(* Schneider Machine Expert - Basic project PROJECT, file version 2.9.0.0 *)
(* ProjectInformations: Name=New project *)

HARDWARE
  Cpu 0: TM221CE16R
  EthernetConfiguration: NetworkName=M221, IpAllocationMode=FixedAddress, IpAddress=0.0.0.0, SubnetMask=0.0.0.0
  SerialLineConfiguration: Baud=Baud19200, Parity=ParityEven, DataBits=DataBits8, StopBits=StopBits1, PhysicalMedium=PhysicalMediumRs485, TransmissionMode=TransmissionModeModbusRtu, SlaveId=1, Addressing=SlaveAddressing
  MastTask: UsePeriodScanMode=false, PeriodScan=100
  FastTask: Period=255
  CpuBehavior: StartingMode=StartAsPreviousState, AutoSaveRamOnEeprom=true, WatchdogPeriod=250

SYMBOLS  (address, symbol, comment, settings)
  %M0         "START"
  %M1         "STOP N RESET"
  %M2         "END CYCLE"
  %M3         "END A"
  %M4         "END B"
  %M10        "BT_START"
  %M11        "BT_RESET"
  %M12        "LAMP IND"
  %M13        "ST VALVE A"
  %M14        "ST VALVE B"
  %M15        "ST VALVE C"
  %M16        "ST AGITATOR"
  %M17        "ST HEATER"
  %M18        "ALARM"
  %S6       SB_TB1S  "Time base of 1 s generated by an internal clock"
  %TM0        "TIMER A"  [Preset=5, Base=OneSecond]
  %TM1        "TIMER B"  [Preset=10, Base=OneSecond]
  %C0         "COUNTER"  [Preset=2]
  %SC0        "COUNTER"
  %I0.0       "START"
  %I0.1       "STOP"
  %I0.2       "SENSOR TINGGI"
  %I0.3       "SENSOR SUHU"
  %Q0.0       "LAMP_INDIKATOR"
  %Q0.1       "VALVE A"
  %Q0.2       "VALVE B"
  %Q0.3       "AGITATOR"
  %Q0.4       "HEATER"
  %Q0.5       "DRAIN VALVE"

POU New POU
  (* SectionNumber=1 *)

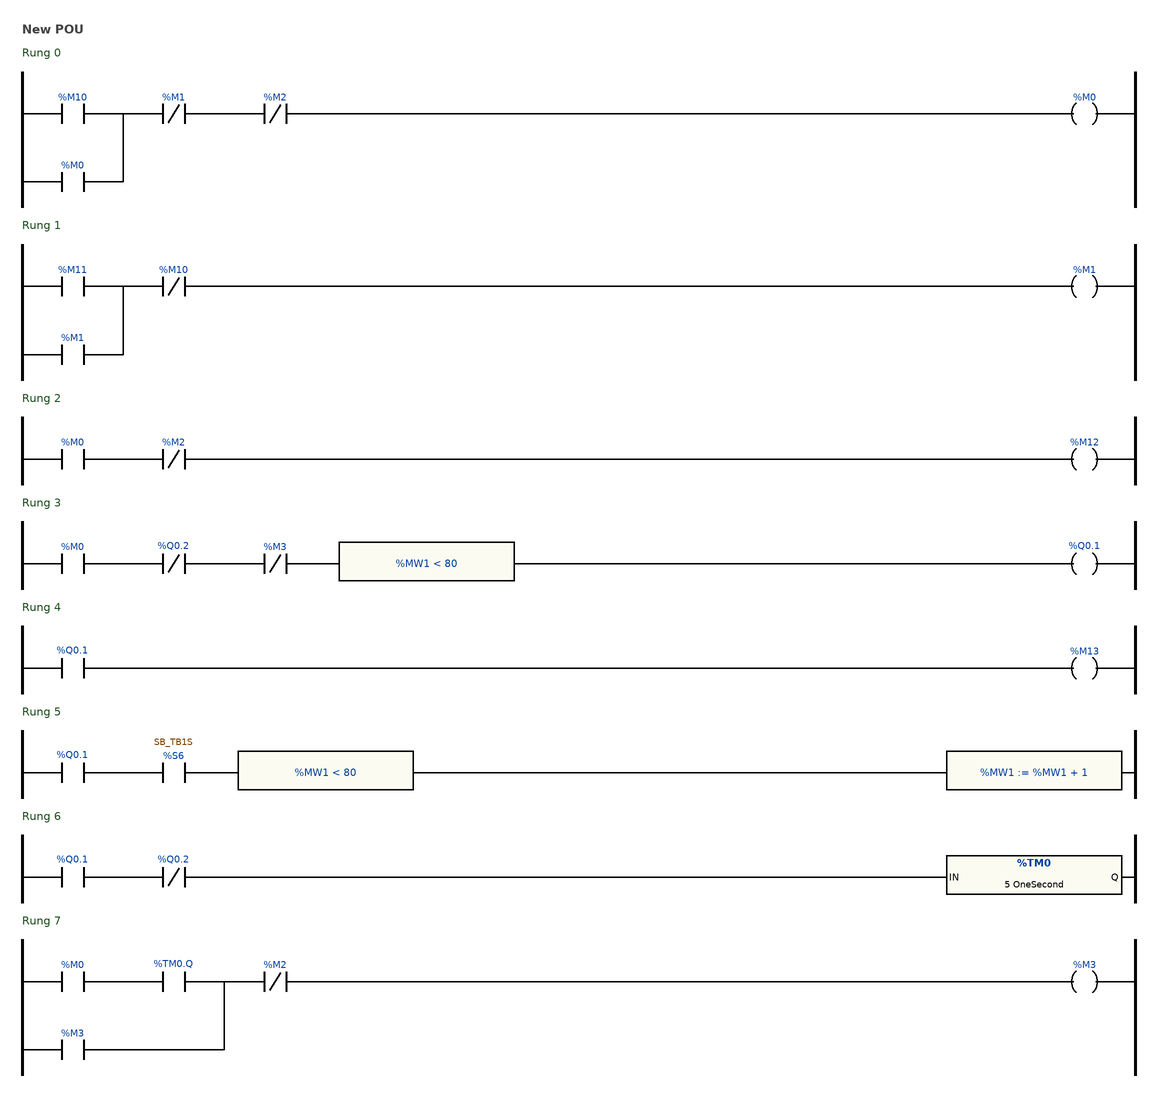

// Rung 0
  LD %M10
  OR %M0
  ANDN %M1
  ANDN %M2
  ST %M0
  // as ST:
  //   %M0 := (%M10 OR %M0) AND NOT %M1 AND NOT %M2;

// Rung 1
  LD %M11
  OR %M1
  ANDN %M10
  ST %M1
  // as ST:
  //   %M1 := (%M11 OR %M1) AND NOT %M10;

// Rung 2
  LD %M0
  ANDN %M2
  ST %M12
  // as ST:
  //   %M12 := %M0 AND NOT %M2;

// Rung 3
  LD %M0
  ANDN %Q0.2
  ANDN %M3
  AND [ %MW1 < 80 ]
  ST %Q0.1
  // as ST:
  //   %Q0.1 := %M0 AND NOT %Q0.2 AND NOT %M3 AND %MW1 < 80;

// Rung 4
  LD %Q0.1
  ST %M13
  // as ST:
  //   %M13 := %Q0.1;

// Rung 5
  LD %Q0.1
  AND %S6                 (* SB_TB1S *)
  AND [ %MW1 < 80 ]
  [ %MW1 := %MW1 + 1 ]
  // as ST:
  //   IF %Q0.1 AND SB_TB1S AND %MW1 < 80 THEN %MW1 := %MW1 + 1; END_IF;

// Rung 6
  BLK %TM0
  LD %Q0.1
  ANDN %Q0.2
  IN
  END_BLK
  // as ST:
  //   %TM0(IN := %Q0.1 AND NOT %Q0.2);

// Rung 7
  LD %M0
  AND %TM0.Q
  OR %M3
  ANDN %M2
  ST %M3
  // as ST:
  //   %M3 := (%M0 AND %TM0.Q OR %M3) AND NOT %M2;

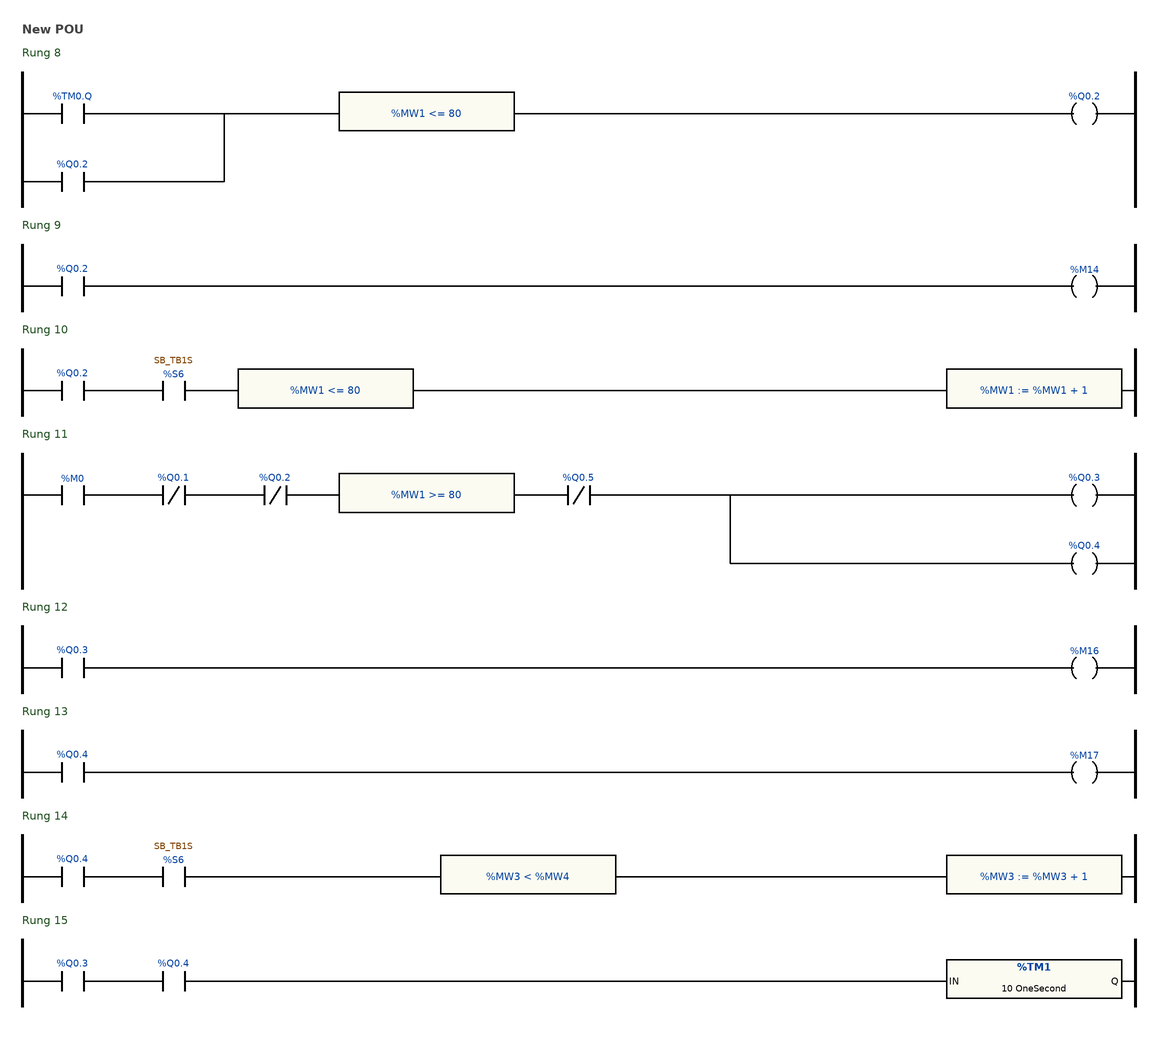

// Rung 8
  LD %TM0.Q
  OR %Q0.2
  AND [ %MW1 <= 80 ]
  ST %Q0.2
  // as ST:
  //   %Q0.2 := (%TM0.Q OR %Q0.2) AND %MW1 <= 80;

// Rung 9
  LD %Q0.2
  ST %M14
  // as ST:
  //   %M14 := %Q0.2;

// Rung 10
  LD %Q0.2
  AND %S6                 (* SB_TB1S *)
  AND [ %MW1 <= 80 ]
  [ %MW1 := %MW1 + 1 ]
  // as ST:
  //   IF %Q0.2 AND SB_TB1S AND %MW1 <= 80 THEN %MW1 := %MW1 + 1; END_IF;

// Rung 11
  LD %M0
  ANDN %Q0.1
  ANDN %Q0.2
  AND [ %MW1 >= 80 ]
  ANDN %Q0.5
  ST %Q0.3
  ST %Q0.4
  // as ST:
  //   %Q0.3 := %M0 AND NOT %Q0.1 AND NOT %Q0.2 AND %MW1 >= 80 AND NOT %Q0.5;
  //   %Q0.4 := %M0 AND NOT %Q0.1 AND NOT %Q0.2 AND %MW1 >= 80 AND NOT %Q0.5;

// Rung 12
  LD %Q0.3
  ST %M16
  // as ST:
  //   %M16 := %Q0.3;

// Rung 13
  LD %Q0.4
  ST %M17
  // as ST:
  //   %M17 := %Q0.4;

// Rung 14
  LD %Q0.4
  AND %S6                 (* SB_TB1S *)
  AND [ %MW3 < %MW4 ]
  [ %MW3 := %MW3 + 1 ]
  // as ST:
  //   IF %Q0.4 AND SB_TB1S AND %MW3 < %MW4 THEN %MW3 := %MW3 + 1; END_IF;

// Rung 15
  BLK %TM1
  LD %Q0.3
  AND %Q0.4
  IN
  END_BLK
  // as ST:
  //   %TM1(IN := %Q0.3 AND %Q0.4);

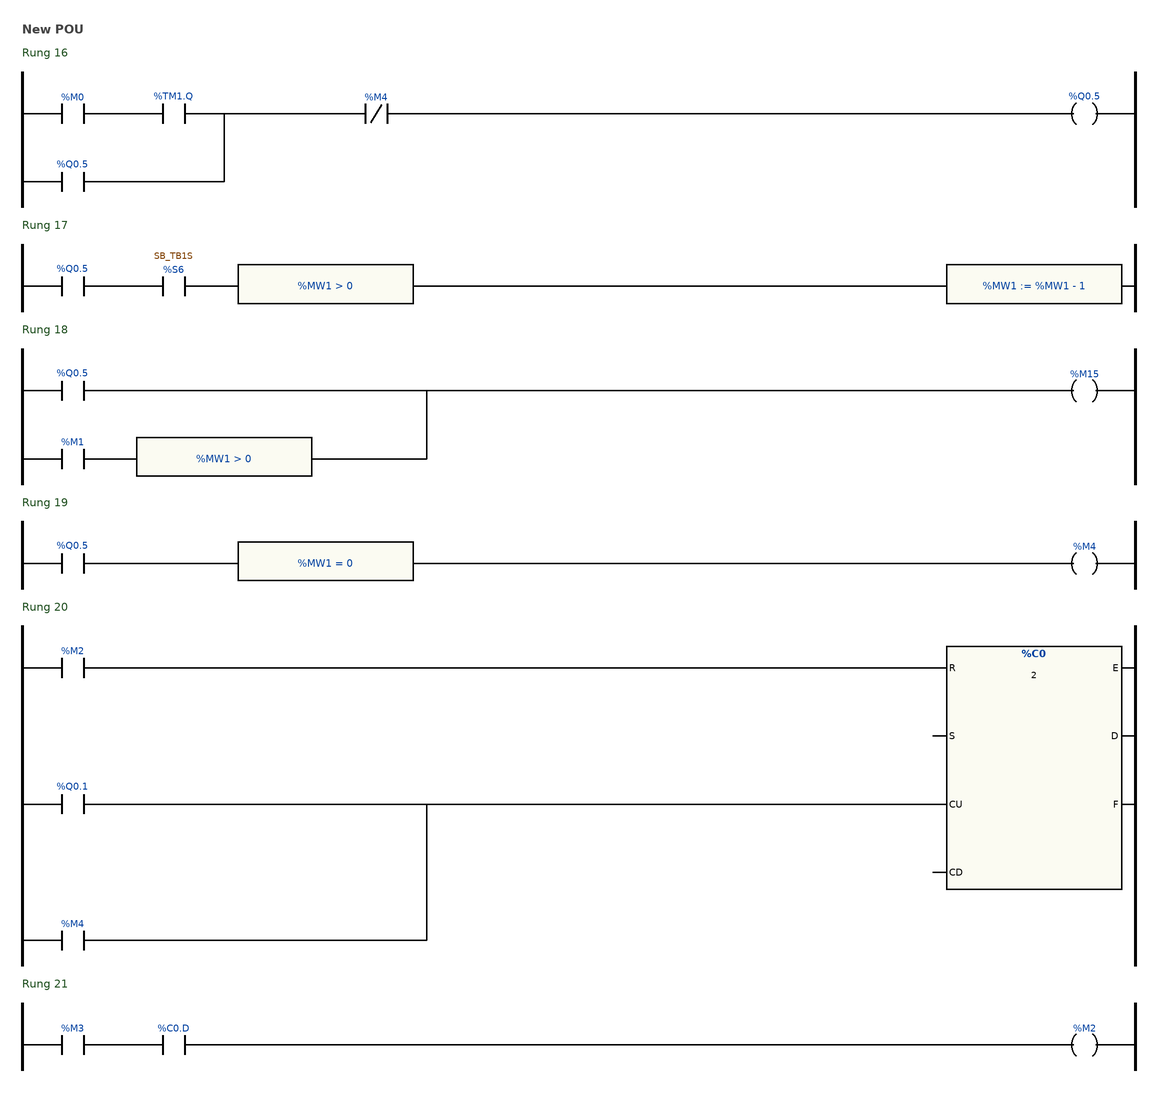

// Rung 16
  LD %M0
  AND %TM1.Q
  OR %Q0.5
  ANDN %M4
  ST %Q0.5
  // as ST:
  //   %Q0.5 := (%M0 AND %TM1.Q OR %Q0.5) AND NOT %M4;

// Rung 17
  LD %Q0.5
  AND %S6                 (* SB_TB1S *)
  AND [ %MW1 > 0 ]
  [ %MW1 := %MW1 - 1 ]
  // as ST:
  //   IF %Q0.5 AND SB_TB1S AND %MW1 > 0 THEN %MW1 := %MW1 - 1; END_IF;

// Rung 18
  LD %Q0.5
  OR( %M1
  AND [ %MW1 > 0 ]
  )
  ST %M15
  // as ST:
  //   %M15 := %Q0.5 OR %M1 AND %MW1 > 0;

// Rung 19
  LD %Q0.5
  AND [ %MW1 = 0 ]
  ST %M4
  // as ST:
  //   %M4 := %Q0.5 AND %MW1 = 0;

// Rung 20
  BLK %C0
  LD %M2
  R
  LD %Q0.1
  OR %M4
  CU
  END_BLK
  // as ST:
  //   %C0(R := %M2, CU := %Q0.1 OR %M4);

// Rung 21
  LD %M3
  AND %C0.D
  ST %M2
  // as ST:
  //   %M2 := %M3 AND %C0.D;

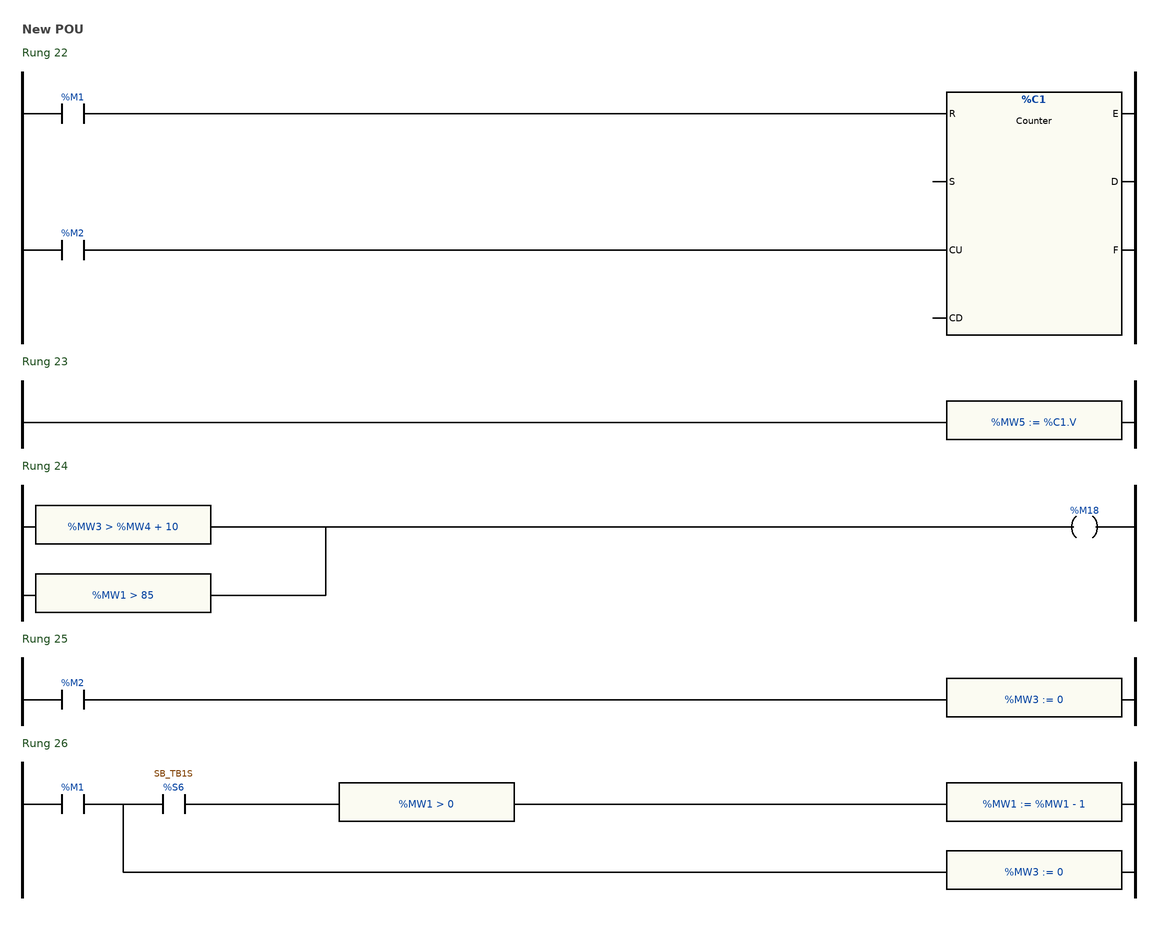

// Rung 22
  BLK %C1
  LD %M1
  R
  LD %M2
  CU
  END_BLK
  // as ST:
  //   %C1(R := %M1, CU := %M2);

// Rung 23
  LD 1
  [ %MW5 := %C1.V ]
  // as ST:
  //   %MW5 := %C1.V;

// Rung 24
  LD 1
  AND [%MW3 > %MW4 + 10]
  OR [ %MW1 > 85 ]
  ST %M18
  // as ST:
  //   %M18 := %MW3 > %MW4 + 10 OR %MW1 > 85;

// Rung 25
  LD %M2
  [ %MW3 := 0 ]
  // as ST:
  //   IF %M2 THEN %MW3 := 0; END_IF;

// Rung 26
  LD %M1
  MPS
  AND %S6                 (* SB_TB1S *)
  AND [ %MW1 > 0 ]
  [ %MW1 := %MW1 - 1 ]
  MPP
  [ %MW3 := 0 ]
  // as ST:
  //   IF %M1 AND SB_TB1S AND %MW1 > 0 THEN %MW1 := %MW1 - 1; END_IF;
  //   IF %M1 THEN %MW3 := 0; END_IF;
